Universal Robots URScript: T015_codellama_34b-instruct-q4_K_M_baseline_rep1.urscript

def program():
    # Home the robot
    movej(p[0.0, 0.0, 0.0, 0.0, 0.0, 0.0], a=350.0, v=350.0)

    # Move above the marking surface
    movel(p[0.0, 0.0, 0.35, 0.0, 0.0, 0.0], a=300.0, v_lead=300.0)

    # Descend
